(* IEC 61131-3 sources: StewartPlatform/Class/SdiasSafetyManagerFSoE (part 2) *)

              LastSDO.ResponseArrived := TRUE;
            else
              LogError("(SdiasSafetyManagerFSoE::ClassState::NewInst) SDO response arrived when no response was expected");
            end_if;
          end_if;
        else
          LogError("(SdiasSafetyManagerFSoE::ClassSvr::NewInst) SDO transfer failed");
        end_if;
      else
        LogError("(SdiasSafetyManagerFSoE::ClassSvr::NewInst) Received invalid SDO response");
      end_if;

//**********************************************************************************************************************************************************
    _BUS_IF_DATA_POINTER_AVAILABLE:
      // does nothing in the FSoE version
      ret_code := READY;

//**********************************************************************************************************************************************************
    _BUS_IF_RESET_DETECTED:
      // don't overwrite other errors
      if SafetyState = _SafetyClassOK then
        SafetyState := _LostPowerSupply;
      end_if;

      // check if module is requred
      MyPara.uiCmd     := _BUS_IF_GET_REQUIRED_SETTING;
      ToBusInterface.NewInst(pPara:=#MyPara, pResult:=#MyResult);
      if MyResult.aData[0]$t_BusIFRetvalErrorcode = _BUS_IF_RETVAL_OK then
        // if it's required => set required error
        if MyResult.aData[4] then

          MyPara.uiCmd := _BUS_IF_SET_REQUIRED_ERROR;
          ToBusInterface.NewInst(#MyPara, #MyResult);
        end_if;
      end_if;

      // drop config of connected modules

      // initialize the message for the periphery
      MyPara.uiCmd := SDIAS_SET_CLASS_STATE;
      MyPara.aPara[1] := 0;// no device ID
      MyPara.aPara[0] := _NoHardware$DINT;

      // tell the connected IO module objects
      if MaxPlace <> SDIAS_SAFETY_INVALID_MAX_PLACE then
        pSafetyModuleInfo := #aSafetyModuleInfo[0];

        for i := 0 to MaxPlace do
          if pSafetyModuleInfo^.pThis then
            pSafetyModuleInfo^.pThis^.NewInst(#MyPara, #MyResult);
          end_if;

          pSafetyModuleInfo += sizeof(t_SdiasSafetyModuleInfo);
        end_for;
      end_if;

      // tell the hbg (if available)
      if sHBG.pThis then
        sHBG.pThis^.NewInst(#MyPara, #MyResult);
      end_if;

//**********************************************************************************************************************************************************
    _BUS_IF_RESET_GONE_DETECTED:
      if SafetyState = _LostPowerSupply then

        // get safety and serial numbers of connected modules
        bUpdateModuleConfig := TRUE;

        // refetch IDs of connected modules
        eCheckIDSSW := _Wait4Idle;

        SafetyState := _SafetyClassOK;
      end_if;

//**********************************************************************************************************************************************************

    CMD_GET_HARDWARE_DIAGNOSIS:
      //Returns module info
      ret_code := ERROR;
      pResult^.aData[0]$t_HWCGetHardwareDiagnosisOut.retcode := _HWC_RETVAL_ERROR;

      pStr_HWTRequested := pPara^.aPara[0]$t_HWCGetHardwareDiagnosisIn.pStr_HardewareTreeEntry;

      tmpplace := (pStr_HWTRequested+pPara^.aPara[0]$t_HWCGetHardwareDiagnosisIn.us_current_index)^$USINT;

      //Check if pointer is valid
      if aSafetyModuleInfo[tmpplace].pThis then

        // Set Offline Device ID
        pResult^.aData[0]$t_HWCGetHardwareDiagnosisOut.ud_DeviceID := (aSafetyModuleInfo[tmpplace].usExpectedDeviceID AND 2#00111000 ) shr 3;   // Bit 3-5 Modul typ
        pResult^.aData[0]$t_HWCGetHardwareDiagnosisOut.ud_Variante :=  aSafetyModuleInfo[tmpplace].usExpectedDeviceID AND 2#00000111;  // Bit 0-2 Submodul typ

        if aModuleIDs[tmpplace] = aSafetyModuleInfo[tmpplace].usExpectedDeviceID then

          ret_code := READY;
          pResult^.aData$t_HWCGetHardwareDiagnosisOut.retcode := _HWC_RETVAL_OK;

          pResult^.aData[0]$t_HWCGetHardwareDiagnosisOut.ud_DeviceID  := (aModuleIDs[tmpplace] AND 2#00111000 ) shr 3;  // Bit 3-5 Modul typ
          pResult^.aData[0]$t_HWCGetHardwareDiagnosisOut.ud_Variante  :=  aModuleIDs[tmpplace] AND 2#00000111; // // Bit 0-2 Submodul typ
          pResult^.aData[0]$t_HWCGetHardwareDiagnosisOut.ud_Place     := tmpplace;

          // Get Serialno ---------------------------------------------------------------------------------------------
          _memcpy(ptr1 := #a_SerialNo[0]
                , ptr2 := #sSafetySerNrs.aSerialNumbers[tmpplace]
                , cntr := sizeof(sSafetySerNrs.aSerialNumbers[tmpplace]) );

          a_SerialNo[sizeof(sSafetySerNrs.aSerialNumbers[tmpplace])] := 0;  // 0 Terminierung

          pResult^.aData[0]$t_HWCGetHardwareDiagnosisOut.pStr_SerialNo := #a_SerialNo[0];

          pResult^.aData[0]$t_HWCGetHardwareDiagnosisOut.hd_SafetyNumber  := sSafetySerNrs.aSafetyNumbers[tmpplace];

        elsif aModuleIDs[tmpplace] <> SDIAS_SAFETY_INVALID_DEVICE_ID then
          pResult^.aData$t_HWCGetHardwareDiagnosisOut.retcode := _HWC_RETVAL_ERROR_WRONG_HARDWARE;
        else
          pResult^.aData$t_HWCGetHardwareDiagnosisOut.retcode := _HWC_RETVAL_ERROR_NO_HARDWARE;
        end_if;

      else
        pResult^.aData[0]$t_HWCGetHardwareDiagnosisOut.retcode := _HWC_RETVAL_ERROR_SDIAS_MODULE_NOT_FOUND;
      end_if;

//**********************************************************************************************************************************************************
    CMD_GET_HARDWARE_TREE_ENTRY:
      //Returns module info

      ret_code := ERROR;
      pResult^.aData[0]$t_HWCGetHardwareTreeEntryOut.retcode := _HWC_RETVAL_ERROR;

      pStr_HWTreeEntry := pPara^.aPara[0]$t_HWCGetHardwareTreeEntryIn.pStr_LastHardewareTreeEntry;

      //First HWT Path
      if (pStr_HWTreeEntry + pStr_HWTreeEntry$^UINT^)^ <> HWT_ESCAPE_INTERNALBUS_SDIAS_SAFETY then  // + 1 for Byte length -1 for 2nd last element of string

        if aSafetyModuleInfo[0].pThis then

          _memcpy(ptr1 := #a_HWTEntryStr[0]
                , ptr2 := pPara^.aPara[0]$t_HWCGetHardwareTreeEntryIn.pStr_LastHardewareTreeEntry
                , cntr := pPara^.aPara[0]$t_HWCGetHardwareTreeEntryIn.pStr_LastHardewareTreeEntry$^UINT^ +2 );  // +2 2 Byte Strlength is not included in the stringlength

          // Add escape sequence
          a_HWTEntryStr[0]$UINT += 1;
          a_HWTEntryStr[a_HWTEntryStr[0]$UINT+1] := HWT_ESCAPE_INTERNALBUS_SDIAS_SAFETY;

          // Add Place
          a_HWTEntryStr[0]$UINT += 1;
          a_HWTEntryStr[a_HWTEntryStr[0]$UINT+1] := 0;

          //Return Hardware Tree Entry and set return codes
          pResult^.aData[0]$t_HWCGetHardwareTreeEntryOut.pStr_NextHardewareTreeEntry := #a_HWTEntryStr[0];

          pResult^.aData[0]$t_HWCGetHardwareTreeEntryOut.retcode := _HWC_RETVAL_OK_HWTSTR_RETURNED;
          ret_code := READY;

        else
          pResult^.aData[0]$t_HWCGetHardwareTreeEntryOut.retcode := _HWC_RETVAL_ERROR_SDIAS_MODULE_NOT_FOUND;
        end_if;

      //search next module
      else

        usNextPlace := (pStr_HWTreeEntry  + pPara^.aPara[0]$t_HWCGetHardwareTreeEntryIn.us_current_index)^$USINT+1;

        if usNextPlace <= SDIAS_SAFETY_MAX_PLACE_NR &
           aSafetyModuleInfo[usNextPlace].pThis then

          _memcpy(ptr1 := #a_HWTEntryStr[0]
                , ptr2 := pPara^.aPara[0]$t_HWCGetHardwareTreeEntryIn.pStr_LastHardewareTreeEntry
                , cntr := pPara^.aPara[0]$t_HWCGetHardwareTreeEntryIn.pStr_LastHardewareTreeEntry$^UINT^ +2 );  // +2 2 Byte Strlength is not included in the stringlength

          // Set new Place
          a_HWTEntryStr[a_HWTEntryStr[0]$UINT + 1] := usNextPlace;

          pResult^.aData[0]$t_HWCGetHardwareTreeEntryOut.pStr_NextHardewareTreeEntry := #a_HWTEntryStr[0];

          //Return Hardware Tree Entry and set return codes
          pResult^.aData[0]$t_HWCGetHardwareTreeEntryOut.retcode := _HWC_RETVAL_OK_HWTSTR_RETURNED;
          ret_code := READY;

        else
          ret_code := READY;
          pResult^.aData$t_HWCGetHardwareTreeEntryOut.retcode := _HWC_RETVAL_OK_END_OF_LIST;
        end_if;
      end_if;

//**********************************************************************************************************************************************************

//*****************************************************************************
//** INTERNAL COMMANDS                                                       **
//*****************************************************************************

//**********************************************************************************************************************************************************
    CMD_SM_READ_PDO_SIZE:
      // get the size of the PDO
      LastSDO.Command := _BUS_IF_READ_VIA_SDO;
      LastSDO.Offset  := SBF_OFFSET_SPDO_LENGTH;
      LastSDO.Length  := sizeof(UINT);

      MyPara.uiCmd    := LastSDO.Command$UINT;
      MyPara.aPara[0] := LastSDO.Offset;
      MyPara.aPara[1] := LastSDO.Length;
      ret_code := ToBusInterface.NewInst(#MyPara, #MyResult);

//**********************************************************************************************************************************************************
  else
    ret_code := SafetyBaseFSoE::NewInst(pPara, pResult);
//**********************************************************************************************************************************************************
	END_CASE;

END_FUNCTION

FUNCTION VIRTUAL SdiasSafetyManagerFSoE::ShowProjectRevision

  ProjectNameStr.WriteDataOff(udLen:=PrjNameStrLen + 1, udOff:=0, pData:=pPrjNameStr);

  ProjectRevisionStr.WriteDataOff(udLen:=PrjRevStrLen + 1, udOff:=0, pData:=pPrjRevStr);

END_FUNCTION

FUNCTION VIRTUAL SdiasSafetyManagerFSoE::InitSafeModule
	VAR_OUTPUT
		sd_retval 	: DINT;
	END_VAR

  // allocate memory for finding unsafe-IO-Servers
  // in first place we allocate 512 byte for our blocked transfers
  p_BlockedTransferMemory := ToStdLib.Malloc( size := SBF_CONFIG_MEMORY_BLOCK_SIZE );
  IF p_BlockedTransferMemory <> NIL THEN
    ud_BlockedTransferMemorySize := SBF_CONFIG_MEMORY_BLOCK_SIZE;
  ELSE
    SafetyState := _MemAllocFailed;
    sd_retval := -100;
    return;
  END_IF;

  // if there is a safety manager to gather the configuration
  if pSafetyManagerThis then
    // allocate memory for gathering configuration information => in first place we allocate 512 byte
    pConfigMem := ToStdLib.Malloc( size := SBF_CONFIG_MEMORY_BLOCK_SIZE );
    IF pConfigMem <> NIL THEN
      ConfigMemSize := SBF_CONFIG_MEMORY_BLOCK_SIZE;
      ConfigMemSizeUsed := 4;
    ELSE
      SafetyState := _MemAllocFailed;
      sd_retval := -100;
      return;
    END_IF;
  end_if;

END_FUNCTION

FUNCTION VIRTUAL GLOBAL SdiasSafetyManagerFSoE::CanOut::NewInst
	VAR_INPUT
		pPara 	: ^CmdStruct;
		pResult 	: ^results;
	END_VAR
	VAR_OUTPUT
		ret_code 	: iprStates;
	END_VAR
  VAR
  	tempCmd         : CmdStruct;
    _result         : results;
  END_VAR

	CASE pPara^.uiCmd OF
//**********************************************************************************************************************************************************
		SDIAS_SAFETY_LOGIN_HBG:
      // check parameters
      if pPara^.aPara[0] & pPara^.aPara[1] then

        sHBG.pThis               := pPara^.aPara[0]$pVirtualBase;
        sHBG.usExpectedDeviceID  := pPara^.aPara[1]$USINT;
        sHBG.sdRequired          := pPara^.aPara[2];
        sHBG.pIOStates           := pPara^.aPara[3]$^HDINT;

        // if leds/hgb not added so far, add them
        if StateBytesUsed = 0 then
          StateBitsUsed := (sizeof(t_LedAndIOStates.biLEDs) + sizeof(t_LedAndIOStates.HBGInputs)) * 8;
          // refresh state bytes used value
          StateBytesUsed := ((StateBitsUsed-1) / 8) + 1;
        end_if;

        if sHBG.sdRequired & (b_AnyModuleRequired = FALSE) then
          b_AnyModuleRequired := TRUE;
          // if any access is required => the businterface is also required
          tempCmd.uiCmd := _BUS_IF_SET_REQUIRED;
          ToBusInterface.NewInst(pPara:=#tempCmd, pResult:=#_result);
          if _result.aData[0]$t_BusIFRetvalErrorcode <> _BUS_IF_RETVAL_OK then
            LogError("(SdiasSafetyManagerFSoE::CanOut::NewInst) Failed to set the BusInterface to required");
          end_if;
        end_if;
      else
        ret_code := ERROR;
      end_if;
//**********************************************************************************************************************************************************
	END_CASE;

	ret_code := READY;

END_FUNCTION

FUNCTION VIRTUAL SdiasSafetyManagerFSoE::GetConfiguration
  VAR
  	pHelp                 : ^void;
    SizeToGo              : UINT;
    ActSize               : UINT;
    ActAddr               : HDINT;
    SDOReqBuf             : SDORequReadConfig;
    SDORspBuf             : ARRAY [0..SBF_SDO_MAX_LENGTH-1] OF USINT;
    pRspBuf               : ^SDORespReadConfig;
    i                     : DINT;
    pSafetyModuleInfo     : ^t_SdiasSafetyModuleInfo;
		MyPara 	              : CmdStruct;
		MyResult              : Results;
  END_VAR

  //initialize header-data for request

  //calculate length without crc
  SDOReqBuf.StdHeader.Len := sizeof(SDORequReadConfig) - sizeof(SDOHeader.StdHeader.CRC);

  //type
  SDOReqBuf.StdHeader.Typ := SDO_STD;

  //command for reading config data
  SDOReqBuf.StdHeader.Cmd := SBF_SDO_COMMAND_READ;

  // read the complete 256 Bytes of safety and serial number info
  pHelp    := #sSafetySerNrs;
  SizeToGo := sizeof(sSafetySerNrs);
  pRspBuf  := (#SDORspBuf)$^SDORespReadConfig;
  ActAddr  := SBF_SDO_ADDRESS_SER_NR_DATA;

  while SizeToGo do
    if SizeToGo > SDIAS_SAFTEY_SDO_MAX_DATA_PER_PAKET then
      ActSize := SDIAS_SAFTEY_SDO_MAX_DATA_PER_PAKET;
    else
      ActSize := SizeToGo;
    end_if;

    if SDOReadCfgRequ(p_SDORequestBuffer  := #SDOReqBuf,
                      p_SDOResponseBuffer := pRspBuf,
                      ud_Address          := ActAddr,
                      us_Length           := ActSize$USINT,
                      b_UseCache          := FALSE) then
      LogError("(SdiasSafetyManagerFSoE::GetConfiguration) Failed to get safety and serial numbers of the IO modules");
      return;
    else
      _memcpy(ptr1:=pHelp, ptr2:=#pRspBuf^.ud_Data, cntr:=ActSize);
    end_if;

    SizeToGo  -= ActSize;
    ActAddr   += ActSize;
    pHelp     += ActSize;
  end_while;

  // only available for IOs, not the HBG
  if MaxPlace <> SDIAS_SAFETY_INVALID_MAX_PLACE then
    // always the same command
    MyPara.uiCmd := SDIAS_SET_NUMBERS;

    pSafetyModuleInfo := #aSafetyModuleInfo[0];
    for i := 0 to MaxPlace$DINT do
      // safety number
      MyPara.aPara[0] := (sSafetySerNrs.aSafetyNumbers[i])$DINT;

      // pointer to serial number string
      MyPara.aPara[1] := (#sSafetySerNrs.aSerialNumbers[i][0])$DINT;

      pSafetyModuleInfo^.pThis^.NewInst(#MyPara, #MyResult);

      pSafetyModuleInfo += sizeof(t_SdiasSafetyModuleInfo);
    end_for;
  end_if;

END_FUNCTION

FUNCTION VIRTUAL GLOBAL SdiasSafetyManagerFSoE::DisconnectEvent
  VAR
  	i                 : UDINT;
    pSafetyModuleInfo : ^t_SdiasSafetyModuleInfo;
		MyPara 	          : CmdStruct;
		MyResult          : Results;
  END_VAR

  SafetyBaseFSoE::DisconnectEvent();

  // initialize the message for the periphery
  MyPara.uiCmd := SDIAS_SET_CLASS_STATE;
  MyPara.aPara[1] := 0;// no device ID
  MyPara.aPara[0] := _NoHardware$DINT;

  // tell the connected IO module objects
  if MaxPlace <> SDIAS_SAFETY_INVALID_MAX_PLACE then
    pSafetyModuleInfo := #aSafetyModuleInfo[0];

    for i := 0 to MaxPlace do
      if pSafetyModuleInfo^.pThis then
        pSafetyModuleInfo^.pThis^.NewInst(#MyPara, #MyResult);
      end_if;

      pSafetyModuleInfo += sizeof(t_SdiasSafetyModuleInfo);
    end_for;
  end_if;

  // tell the hbg (if available)
  if sHBG.pThis then
    sHBG.pThis^.NewInst(#MyPara, #MyResult);
  end_if;

  // clear the strings
  ProjectNameStr.Clear();
  ProjectRevisionStr.Clear();

END_FUNCTION

FUNCTION VIRTUAL SdiasSafetyManagerFSoE::SetSafetyState
	VAR_INPUT
		NewState 	: SafetyConfigStateType;
	END_VAR
  VAR
		MyPara 	  : CmdStruct;
		MyResult	: results;
  END_VAR

  // use it locally
  SafetyState := NewState;

  // tell the outer class
  MyPara.uiCmd := SDIAS_SET_SAFETY_STATE;
  MyPara.aPara[0] := NewState$DINT;
  ToBusInterface.NewInst(#MyPara, #MyResult);

END_FUNCTION

FUNCTION VIRTUAL GLOBAL SdiasSafetyManagerFSoE::CyWork
	VAR_INPUT
		EAX 	: UDINT;
	END_VAR
	VAR_OUTPUT
		state (EAX) 	: UDINT;
	END_VAR
  VAR
		MyPara 	          : CmdStruct;
		MyResult          : Results;
    TmpRetCode        : iprStates;
  END_VAR

  // if the initialisiation has been finished and there is an object for the hbg check if it's has been connected or disconnected
  if Online then

    case eCheckIDSSW of
  //**********************************************************************************************************************************************************
      _Nothing:
        if sHBG.pThis then
          // check for a can connect event
          if CanActive > OldCanActive then
            // if we're already idle => get it on
            if eResponseState = _idle then
              eCheckIDSSW := _GetIDs;
            else
              // otherwise, wait for it (need to remember the connect event)
              eCheckIDSSW := _Wait4Idle;
            end_if;

          // check for a can disconnect event
          elsif CanActive < OldCanActive then
            if sHBG.sdRequired then
              // if it's required => required error
              MyPara.uiCmd := _BUS_IF_SET_REQUIRED_ERROR;
              ToBusInterface.NewInst(#MyPara, #MyResult);
            else
              // otherwise show that it has been disconnected
              MyPara.uiCmd := SDIAS_SET_CLASS_STATE;
              MyPara.aPara[1] := 0;// no device ID
              MyPara.aPara[0] := _NoHardware$DINT;
              sHBG.pThis^.NewInst(#MyPara, #MyResult);
            end_if;
          end_if;
          OldCanActive := CanActive;
        end_if;

  //**********************************************************************************************************************************************************
      _Wait4Idle:
        if eResponseState = _idle then
          eCheckIDSSW := _GetIDs;
        end_if;

  //**********************************************************************************************************************************************************
      _GetIDs:
        case eResponseState of
        //*****************************************************
          _idle:
            LastSDO.Command := _BUS_IF_READ_VIA_SDO;
            LastSDO.Offset  := SBF_OFFSET_IO_MODULE_IDS;
            LastSDO.Length  := sizeof(t_ModuleIDs);

            MyPara.uiCmd    := LastSDO.Command$UINT;
            MyPara.aPara[0] := LastSDO.Offset;
            MyPara.aPara[1] := LastSDO.Length;
            TmpRetcode := ToBusInterface.NewInst(#MyPara, #MyResult);
            if TmpRetcode = READY then
              SDOTimeMark  := ops.tAbsolute;
              eResponseState:= _wait;
            elsif TmpRetcode = ERROR then
              LogError("(SdiasSafetyManagerFSoE::InitModule) Failed to add read SDO for module configuration");
            end_if;
        //*****************************************************
          _wait:
            // wait for response
            if ((ops.tAbsolute - SDOTimeMark) > SDIAS_SAFTEY_SDO_RESPONSE_TIMEOUT) then
              LogError("(SdiasSafetyManagerFSoE::InitModule) SDO Response timeout while waiting for the module configuration");
              eCheckIDSSW := _Nothing;
              eResponseState := _idle;
            end_if;
        //*****************************************************
          _valid:
            eCheckIDSSW := _Nothing;
            eResponseState := _idle;
        //*****************************************************
        end_case;
  //**********************************************************************************************************************************************************
    end_case;
  end_if;

	state := SafetyBaseFSoE::CyWork(0);

END_FUNCTION

FUNCTION VIRTUAL SdiasSafetyManagerFSoE::RefreshAsySrv
  VAR
  	i                 : UDINT;
    pSafetyModuleInfo : ^t_SdiasSafetyModuleInfo;
		MyPara 	          : CmdStruct;
		MyResult          : Results;
    AsyValues         : t_AsyRefresh;
  END_VAR

  // tell the outer class
  MyPara.uiCmd := SDIAS_SET_ASY_STATE;
  AsyValues.QuitComError := QuitComError;
  MyPara.aPara[0] := (#AsyValues)$DINT;
  ToBusInterface.NewInst(#MyPara, #MyResult);

  // tell the connected IO module objects
  if MaxPlace <> SDIAS_SAFETY_INVALID_MAX_PLACE then
    pSafetyModuleInfo := #aSafetyModuleInfo[0];

    for i := 0 to MaxPlace do
      if pSafetyModuleInfo^.pThis then
        pSafetyModuleInfo^.pThis^.NewInst(#MyPara, #MyResult);
      end_if;

      pSafetyModuleInfo += sizeof(t_SdiasSafetyModuleInfo);
    end_for;
  end_if;

END_FUNCTION

FUNCTION VIRTUAL GLOBAL SdiasSafetyManagerFSoE::FastUnsafeOutputs::Write
	VAR_INPUT
		input (EAX) 	: BDINT;
	END_VAR
	VAR_OUTPUT
		result (EAX) 	: BDINT;
	END_VAR
  VAR
  	pUnsafeOutLogin : ^t_FastUnsafeOuts;
  END_VAR

  // if the pointer is valid and we're in the first init run (the firstscan check prevents a crash caused by someone writing on the server during runtime)
	if input & (us_FirstScan < 2) then
    pUnsafeOutLogin := input$^t_FastUnsafeOuts;
    // check if it's the correct usage of the class
    if pUnsafeOutLogin^.Kennung = SDIAS_SAFETY_FAST_UNSAFE_KENNUNG then
      pFastUnsafeOutThis := pUnsafeOutLogin^.pThis;
    end_if;
  end_if;

	result := input;

END_FUNCTION

FUNCTION VIRTUAL GLOBAL SdiasSafetyManagerFSoE::FastUnsafeInputs::Write
	VAR_INPUT
		input (EAX) 	: BDINT;
	END_VAR
	VAR_OUTPUT
		result (EAX) 	: BDINT;
	END_VAR

	FastUnsafeInputs := input;
	result := FastUnsafeInputs;

END_FUNCTION

FUNCTION VIRTUAL SdiasSafetyManagerFSoE::SetRetryCounter
	VAR
    pSafetyModuleInfo : ^t_SdiasSafetyModuleInfo;
		MyPara 	 : CmdStruct;
		MyResult : Results;
    i        :  USINT;
	END_VAR

  if b_RetryCounterAvailable then

    if MaxPlace <> SDIAS_SAFETY_INVALID_MAX_PLACE then
      //Command for new inst call in sdiassafetybase
      MyPara.uiCmd := SDIAS_SET_RETRY_COUNTER;

      //calls newinst method of all safety modules which exists.
      for i := 0 to MaxPlace do
        pSafetyModuleInfo := #aSafetyModuleInfo[i];
        MyPara.aPara[0] := a_RetryCnt[i];
        MyPara.aPara[1] := a_RetryCnt[i+16];  //+16 for retry counter of µC2
        pSafetyModuleInfo^.pThis^.NewInst(#MyPara, #MyResult);
      end_for;
    end_if;
  else
    //Retrycounter not available -> show -1 at servers.
    SafetyRetryCounter := -1; //Not available

    if MaxPlace <> SDIAS_SAFETY_INVALID_MAX_PLACE then
      MyPara.uiCmd := SDIAS_RETRY_COUNTER_NOT_AVAILABLE;
      for i := 0 to MaxPlace do
        pSafetyModuleInfo := #aSafetyModuleInfo[i];
        pSafetyModuleInfo^.pThis^.NewInst(#MyPara, #MyResult);
      end_for;
    end_if;
  end_if;

END_FUNCTION

FUNCTION VIRTUAL GLOBAL SdiasSafetyManagerFSoE::Background
	VAR_INPUT
		EAX 	: UDINT;
	END_VAR
	VAR_OUTPUT
		state (EAX) 	: UDINT;
	END_VAR

  if bUpdateModuleConfig & (eCheckIDSSW = _Nothing) then
    GetConfiguration();
  end_if;

	state := SafetyBaseFSoE::Background(0);

END_FUNCTION

FUNCTION VIRTUAL SdiasSafetyManagerFSoE::BusConfigWrite
	VAR_INPUT
		Offset 	: HDINT;
		Length 	: UINT;
		pData 	: pVoid;
		IsControlAccess 	: BOOL;(* := FALSE *)
	END_VAR
	VAR_OUTPUT
		retcode 	: iprStates;
	END_VAR
  VAR
  	TmpRetcode  : iprStates;
    MyPara      : CmdStruct;
    MyResult    : results;
  END_VAR

  retcode := BUSY;

  case Config.BusConfigSSW of
//**********************************************************************************************************************************************************
    _PrepareAccess:
      Config.RestLength := Length;
      Config.pActData   := pData;

      Config.BusConfigSSW := _StartAccess;

//**********************************************************************************************************************************************************
    _StartAccess:
      if IsControlAccess then
        LastSDO.Command := _BUS_IF_WRITE_VIA_SDO_CTRL;
      else
        LastSDO.Command := _BUS_IF_WRITE_VIA_SDO;
      end_if;

      LastSDO.Offset  := Offset$DINT;
      if Config.RestLength > SDIAS_SAFETY_MAX_SDO_DATA_PER_CYCLE then
        LastSDO.Length  := SDIAS_SAFETY_MAX_SDO_DATA_PER_CYCLE;
      else
        LastSDO.Length  := Config.RestLength;
      end_if;
      LastSDO.ResponseArrived := FALSE;

      MyPara.uiCmd    := LastSDO.Command;
      MyPara.aPara[0] := LastSDO.Offset;
      MyPara.aPara[1] := LastSDO.Length;
      MyPara.aPara[2] := Config.pActData$DINT;
      TmpRetcode := ToBusInterface.NewInst(#MyPara, #MyResult);
      if TmpRetcode = READY then
        Config.SDOTimeMark  := ops.tAbsolute;
        Config.BusConfigSSW := _Wait4Answer;
      elsif TmpRetcode = ERROR then
        retcode := ERROR;
        LogError("(SdiasSafetyManagerFSoE::BusConfigWrite) Failed to add write SDO for module configuration");
      end_if;

//**********************************************************************************************************************************************************
    _Wait4Answer:
      // wait for response

      // check for response
      if LastSDO.ResponseArrived then
        Config.RestLength -= LastSDO.Length;
        Config.pActData   += LastSDO.Length;

        if Config.RestLength = 0 then
          retcode := READY;
          Config.BusConfigSSW := _PrepareAccess;
        end_if;
      elsif ((ops.tAbsolute - Config.SDOTimeMark) > SDIAS_SAFTEY_SDO_RESPONSE_TIMEOUT) then
        LogError("(SdiasSafetyManagerFSoE::BusConfigWrite) SDO Response timeout while waiting for the write response");
        retcode := ERROR;
      end_if;

//**********************************************************************************************************************************************************
  end_case;

END_FUNCTION

FUNCTION VIRTUAL SdiasSafetyManagerFSoE::BusConfigRead
	VAR_INPUT
		Offset 	: HDINT;
		Length 	: UINT;
		pData 	: pVoid;
		IsControlAccess 	: BOOL;(* := FALSE *)
	END_VAR
	VAR_OUTPUT
		retcode 	: iprStates;
	END_VAR
  VAR
  	TmpRetcode  : iprStates;
    MyPara      : CmdStruct;
    MyResult    : results;
  END_VAR

  retcode := BUSY;

  case Config.BusConfigSSW of
//**********************************************************************************************************************************************************
    _PrepareAccess:
      Config.RestLength := Length;
      Config.pActData   := pData;

      Config.BusConfigSSW := _StartAccess;

//**********************************************************************************************************************************************************
    _StartAccess:
      if IsControlAccess then
        LastSDO.Command := _BUS_IF_READ_VIA_SDO_CTRL;
      else
        LastSDO.Command := _BUS_IF_READ_VIA_SDO;
      end_if;

      LastSDO.Offset  := Offset$DINT;
      if Config.RestLength > SDIAS_SAFETY_MAX_SDO_DATA_PER_CYCLE then
        LastSDO.Length  := SDIAS_SAFETY_MAX_SDO_DATA_PER_CYCLE;
      else
        LastSDO.Length  := Config.RestLength;
      end_if;
      LastSDO.ResponseArrived := FALSE;

      MyPara.uiCmd    := LastSDO.Command;
      MyPara.aPara[0] := LastSDO.Offset;
      MyPara.aPara[1] := LastSDO.Length;
      TmpRetcode := ToBusInterface.NewInst(#MyPara, #MyResult);
      if TmpRetcode = READY then
        Config.SDOTimeMark  := ops.tAbsolute;
        Config.BusConfigSSW := _Wait4Answer;
      elsif TmpRetcode = ERROR then
        retcode := ERROR;
        LogError("(SdiasSafetyManagerFSoE::BusConfigRead) Failed to add write SDO for module configuration");
      end_if;

//**********************************************************************************************************************************************************
    _Wait4Answer:
      // wait for response

      // check for response
      if LastSDO.ResponseArrived then
        Config.RestLength -= LastSDO.Length;
        Config.pActData   += LastSDO.Length;

        if Config.RestLength = 0 then
          retcode := READY;
          Config.BusConfigSSW := _PrepareAccess;
        end_if;
      elsif ((ops.tAbsolute - Config.SDOTimeMark) > SDIAS_SAFTEY_SDO_RESPONSE_TIMEOUT) then
        LogError("(SdiasSafetyManagerFSoE::BusConfigRead) SDO Response timeout while waiting for the write response");
        retcode := ERROR;
      end_if;

//**********************************************************************************************************************************************************
  end_case;

END_FUNCTION
